(*
SPDX-FileCopyrightText: © 2026 Oleksandr Tiutyk <trofimich@gmail.com>
SPDX-License-Identifier: MIT
License: https://opensource.org/license/mit
*)

(*!
<summary>Provides constants and helpers for configuration nodes.</summary>
<description>
Supplies canonical boundary values such as EMPTY_NODE for comparisons.
</description>
*)
{attribute 'no_explicit_call' := 'do not call this function block directly'}
PROGRAM ConfigurationNodes
VAR CONSTANT
	//! <summary>Empty configuration node denoting an absent or unassigned node.</summary>
	EMPTY_NODE : CONFIGURATION_NODE := (Handle := 0);
END_VAR
VAR
	{attribute 'hide'}
	_ClassName : STRING := __POUNAME();
END_VAR

(*!
<summary>Returns the program class name for diagnostic reporting.</summary>
*)
{attribute 'monitoring' := 'call'}
PROPERTY ClassName : REFERENCE TO STRING
GET
ClassName REF= _ClassName;
END_GET
END_PROPERTY

(*!
<summary>Returns the library namespace name for diagnostic reporting.</summary>
*)
{attribute 'monitoring' := 'call'}
PROPERTY NamespaceName : REFERENCE TO STRING
GET
NamespaceName REF= CurrentNamespace.Name;
END_GET
END_PROPERTY

END_PROGRAM

(* stored: Version 1.1.0.1
   POU ConfigurationNodes: Id {c9a87487-a25c-431a-a764-27b6c2a15990}, SpecialFunc None
   Property ClassName: Id {eb897fb0-e736-49fd-8507-f399b3e93803}
   Get Get: Id {ede1d259-08dd-4f84-9964-2f27ccf4cb29}
   Property NamespaceName: Id {a0012fb4-1257-49ef-b3c2-7533d3db33bc}
   Get Get: Id {950c767c-0375-4435-8879-bba52c7f142a} *)
